Fanuc KAREL source: kf00083.KL

-- PROVISIONAL review KL for V1013-1; original PC SHA256 9ea9b09afbd3b9ff76bb826eb56cd29a0b80b5adbb0aa4ee6c60c278d750de24
-- Incomplete behavior may be omitted. Consult companion uncertainty JSON. Do not deploy.
PROGRAM KF00083
%NOLOCKGROUP
VAR
  I : INTEGER
  J : INTEGER
  X : REAL
  Y : REAL
  B : BOOLEAN
  C : BOOLEAN
  TXT : STRING[80]
  TXT2 : STRING[80]
  STATUS : INTEGER
-- UNRESOLVED_DECL AI type=002010
-- UNRESOLVED_DECL BI type=002010
-- UNRESOLVED_DECL P type=000102
-- UNRESOLVED_DECL JP type=000199
-- UNRESOLVED_DECL PF type=000101
-- UNRESOLVED_DECL V1 type=000013
-- UNRESOLVED_DECL V2 type=000013
BEGIN
  -- UNRESOLVED_PC offsets 5-26; opcodes 27,27,9C,27,9C,27,9D,76,7E,4A
  -- UNRESOLVED_PC offsets 31-35; opcodes 7F
END KF00083
